(* IEC 61131-3 sources: kns-port-domestic/upstream/plc-process-lib/src/POUs/Devices/FB_AnalogInput, 16 files *)

(* ---- ClassifySignal.method.impl.st ---- *)
IF NOT F_IsFinite(rIn := rIn) THEN
    ClassifySignal := E_AiSignalState.NotFinite;
ELSIF xChannelFault THEN
    ClassifySignal := E_AiSignalState.ChannelFault;
ELSIF stCfgLkg.eInput = E_AiInputType.MilliAmp OR stCfgLkg.eInput = E_AiInputType.Norm420 THEN
    IF stCfgLkg.eInput = E_AiInputType.Norm420 THEN
        rI_mA := GVL_Const.MA_ZERO + GVL_Const.MA_SPAN * rIn;
    ELSE
        rI_mA := rIn;
    END_IF
    IF rI_mA <= GVL_Const.NE43_FAIL_LOW_MA THEN
        ClassifySignal := E_AiSignalState.FailLow;
    ELSIF rI_mA >= GVL_Const.NE43_FAIL_HIGH_MA THEN
        ClassifySignal := E_AiSignalState.FailHigh;
    ELSIF rI_mA < GVL_Const.NE43_MEAS_LOW_MA THEN
        ClassifySignal := E_AiSignalState.UnderRange;
    ELSIF rI_mA > GVL_Const.NE43_MEAS_HIGH_MA THEN
        ClassifySignal := E_AiSignalState.OverRange;
    ELSE
        ClassifySignal := E_AiSignalState.Good;
    END_IF
ELSE
    // Norm01, Eng, Raw: NE 43 не применяется
    ClassifySignal := E_AiSignalState.Good;
END_IF

(* ---- FB_AnalogInput.decl.st ---- *)
// Назначение: аналоговый вход. Сигнал 4–20 мА, нормированный 0–1, инженерные единицы или отсчёты
//             канала → значение в инженерных единицах: достоверность по NAMUR NE 43 с
//             подтверждением tFailDelay и удержанием последнего хорошего значения на время
//             подтверждения, корень с отсечкой малых значений, фильтр первого порядка по реальному
//             шагу времени, уставки HH/H/L/LL (FB_LimitMonitor), подмена значения с ограничением по
//             времени, шесть слотов тревог. Режимы: Auto — измерение, Manual — подмена,
//             OutOfService; Local нет. Наследует FB_DeviceBase: тело — нормативный порядок цикла,
//             шаги обработки сигнала — защищённые методы.
// Автор:      kr0nsch
// Версия:     0.1.0
// Документ:   docs/fb/FB_AnalogInput.md
FUNCTION_BLOCK FB_AnalogInput EXTENDS FB_DeviceBase
VAR_INPUT
    rIn                  : REAL;     // значение канала; смысл — по stCfg.eInput
    xChannelFault        : BOOL;     // диагностика модуля или ошибка обмена (для значений по Modbus)
    xSuppressLimitAlarms : BOOL;     // подавить тревоги уставок по условию (флаги уставок считаются)
END_VAR
VAR_IN_OUT
    stCmd : ST_AnalogInputCmd;       // команды HMI/SCADA (GVL_Hmi.st<TAG>Cmd)
END_VAR
VAR_IN_OUT CONSTANT
    stCfg : ST_AnalogInputCfg;       // параметры (GVL_Persist.st<TAG>Cfg), только чтение
END_VAR
VAR_OUTPUT
    rValue_eu  : REAL;               // значение для логики, инж. ед.
    rValue_pct : REAL;               // значение, % шкалы
    xValid     : BOOL;               // значение пригодно для управления
    xHH        : BOOL;               // верхняя аварийная уставка (после гистерезиса и задержек)
    xH         : BOOL;               // верхняя предупредительная уставка
    xL         : BOOL;               // нижняя предупредительная уставка
    xLL        : BOOL;               // нижняя аварийная уставка
    stSts      : ST_AnalogInputSts;  // состояние для HMI/SCADA
END_VAR
VAR
    stCfgLkg  : ST_AnalogInputCfg;                       // последняя корректная конфигурация (LKG)
    afbLimit  : ARRAY[0..3] OF FB_LimitMonitor;          // уставки, индекс E_AiAlarm.HH, H, L, LL
    fbFail    : FB_Delay;                                // подтверждение отказа сигнала и возврата
    fbOor     : FB_Delay;                                // подтверждение выхода за диапазон и возврата
    fbSubst   : FB_Delay;                                // длительность подмены (tSubstMax)
    eSignal   : E_AiSignalState := E_AiSignalState.Good; // мгновенная классификация сигнала
    xRawFail  : BOOL;                                    // мгновенный отказ сигнала (до подтверждения)
    xFail     : BOOL;                                    // отказ сигнала подтверждён
    xOor      : BOOL;                                    // выход за диапазон подтверждён
    xValueBad : BOOL;                                    // измеренного значения нет: отказ подтверждён
                                                         // или хорошего значения ещё не было
    lrFlt     : LREAL;                                   // состояние фильтра, инж. ед.
    xFltInit  : BOOL := TRUE;                            // фильтр начнётся с текущего значения
    rGood_eu  : REAL;                                    // последнее хорошее значение, инж. ед.
    xHaveGood : BOOL;                                    // хорошее значение было после старта ПЛК или
                                                         // после возврата контроля (OutOfService, Cfg)
    xLowCut   : BOOL;                                    // сработала отсечка малых значений
    xClamped  : BOOL;                                    // значение ограничено шкалой
END_VAR
VAR_TEMP
    eRes       : E_CmdResult;        // результат ProcessMode
    xRawOor    : BOOL;               // мгновенный выход за диапазон (до подтверждения)
    xSupervise : BOOL;               // контроль сигнала: корректная Cfg была, не OutOfService
    xLimOff    : BOOL;               // флаги уставок снять сразу
    xLimSupp   : BOOL;               // подавление тревог уставок
    wLowBits   : WORD;               // младший байт wStatus
    eDevSt     : E_Ne107Status;      // вклад логики устройства в NE 107
END_VAR

(* ---- CallLimit.method.decl.st ---- *)
// Вызов одной уставки FB_LimitMonitor (шаг 7 цикла), результат — флаг уставки xOut. Уставка
// передаётся через VAR_IN_OUT: шаг уставок в теле — один вызов на уставку (AI-1). Внутренний шаг
// устройства: PROTECTED (правило L5 контракта), имя зарезервировано
METHOD PROTECTED CallLimit : BOOL
VAR_INPUT
    rLimValue : REAL;              // контролируемое значение, инж. ед.
    xHigh     : BOOL;              // TRUE — верхняя уставка (HH, H), FALSE — нижняя (L, LL)
    xOff      : BOOL;              // снять флаг сразу (OutOfService, нет Cfg, отказ)
    stLimCfg  : ST_AiLimitCfg;     // параметры уставки (stCfgLkg.astLimit[i])
END_VAR
VAR_IN_OUT
    fbLimit : FB_LimitMonitor;     // уставка afbLimit[i]
END_VAR

(* ---- CheckConfig.method.decl.st ---- *)
// Проверка конфигурации: биты wCfgErr аналогового входа (карта — docs/fb/FB_AnalogInput.md). Только
// считает, ничего не меняет. Сравнения записаны так, чтобы NaN давал ошибку (NOT (x >= a AND x <= b))
METHOD PROTECTED CheckConfig : WORD
VAR_IN_OUT CONSTANT
    stCfgIn : ST_AnalogInputCfg;   // проверяемая конфигурация
END_VAR
VAR
    wErr    : WORD;                // непройденные проверки
    uiIdx   : UINT;                // индекс уставки: HH, H, L, LL
    stLim   : ST_AiLimitCfg;       // копия уставки: короче условия проверок
    xPrev   : BOOL;                // была включённая уставка старше текущей
    rPrevSp : REAL;                // её значение, инж. ед.
    rSpan   : REAL;                // диапазон шкалы, инж. ед.
END_VAR

(* ---- CheckConfig.method.impl.st ---- *)
IF NOT (stCfgIn.eInput = E_AiInputType.MilliAmp OR stCfgIn.eInput = E_AiInputType.Norm420
        OR stCfgIn.eInput = E_AiInputType.Norm01 OR stCfgIn.eInput = E_AiInputType.Eng
        OR stCfgIn.eInput = E_AiInputType.Raw)
THEN
    wErr := wErr OR GVL_Const.AI_CFG_INPUT_TYPE;
END_IF
IF NOT (F_IsFinite(rIn := stCfgIn.rRangeLo_eu) AND F_IsFinite(rIn := stCfgIn.rRangeHi_eu)
        AND stCfgIn.rRangeLo_eu < stCfgIn.rRangeHi_eu)
THEN
    wErr := wErr OR GVL_Const.AI_CFG_RANGE;
END_IF

// Уставки: включённые — в шкале, гистерезис 0 <= h < диапазона, порядок строго LL < L < H < HH
// (обход от HH к LL: каждая следующая включённая строго меньше предыдущей включённой)
rSpan := stCfgIn.rRangeHi_eu - stCfgIn.rRangeLo_eu;
FOR uiIdx := E_AiAlarm.HH TO E_AiAlarm.LL DO
    stLim := stCfgIn.astLimit[uiIdx];
    IF stLim.xEnable THEN
        IF NOT (stLim.rSetpoint_eu >= stCfgIn.rRangeLo_eu AND stLim.rSetpoint_eu <= stCfgIn.rRangeHi_eu) THEN
            wErr := wErr OR GVL_Const.AI_CFG_LIMIT_OUT_OF_RANGE;
        END_IF
        IF NOT (F_IsFinite(rIn := stLim.rHyst_eu) AND stLim.rHyst_eu >= 0.0 AND stLim.rHyst_eu < rSpan) THEN
            wErr := wErr OR GVL_Const.AI_CFG_HYST;
        END_IF
        IF xPrev AND NOT (stLim.rSetpoint_eu < rPrevSp) THEN
            wErr := wErr OR GVL_Const.AI_CFG_LIMIT_ORDER;
        END_IF
        xPrev := TRUE;
        rPrevSp := stLim.rSetpoint_eu;
    END_IF
END_FOR

IF NOT (stCfgIn.rLowCut_pct >= 0.0 AND stCfgIn.rLowCut_pct <= GVL_Const.AI_LOWCUT_MAX_PCT) THEN
    wErr := wErr OR GVL_Const.AI_CFG_LOW_CUT;
END_IF
IF NOT (stCfgIn.eFailValue = E_AiFailValue.HoldLast OR stCfgIn.eFailValue = E_AiFailValue.Substitute)
   OR NOT F_IsFinite(rIn := stCfgIn.rFailValue_eu)
THEN
    wErr := wErr OR GVL_Const.AI_CFG_FAIL_VALUE;
END_IF
IF NOT CheckAlarmCfg(astCfg := stCfgIn.astAlarm) THEN
    wErr := wErr OR GVL_Const.AI_CFG_ALARM;
END_IF
// шкала отсчётов проверяется только у входа Raw: умолчания 0/0 проходят у остальных типов
IF stCfgIn.eInput = E_AiInputType.Raw
   AND NOT (F_IsFinite(rIn := stCfgIn.rRawLo_cnt) AND F_IsFinite(rIn := stCfgIn.rRawHi_cnt)
            AND stCfgIn.rRawLo_cnt < stCfgIn.rRawHi_cnt)
THEN
    wErr := wErr OR GVL_Const.AI_CFG_RAW_RANGE;
END_IF
CheckConfig := wErr;

(* ---- ClassifySignal.method.decl.st ---- *)
// Шаг 6.1 цикла: мгновенная классификация сигнала (до подтверждения tFailDelay). NE 43 — только для
// MilliAmp и Norm420 (I = 4 + 16·rIn); старшинство NotFinite > ChannelFault > FailLow/FailHigh >
// UnderRange/OverRange > Good. Границы 3,6 и 21,0 мА включены в отказ (A-02, сверить с NAMUR NE 43).
// Читает входы rIn, xChannelFault и stCfgLkg; ничего не меняет
METHOD PROTECTED ClassifySignal : E_AiSignalState
VAR
    rI_mA : REAL;   // ток для проверки NE 43, мА
END_VAR

(* ---- ComputeValue.method.decl.st ---- *)
// Шаг 6.3 цикла (LREAL): нормировка по типу входа, корень и отсечка малых значений, инженерные
// единицы, ограничение шкалой, фильтр первого порядка — точная экспонента по реальному шагу времени.
// 4–20 мА (MilliAmp, Norm420): значение не экстраполируется за насыщение NE 43 (3,8 и 20,5 мА, AI-13)
// ltDt (реакция не зависит от цикла). Без расчёта (xCompute = FALSE: нет корректной Cfg, OutOfService,
// отказ сигнала) фильтр стоит. После подтверждённого отказа и после возврата контроля (xRestart) фильтр
// начинается с текущего значения, без «подтягивания» от старого; короткий неподтверждённый провал
// фильтр только замораживает — после него значение продолжается без скачка (AI-12). Хорошее значение
// для удержания запоминается, пока отказ не подтверждён
METHOD PROTECTED ComputeValue
VAR_INPUT
    xCompute : BOOL;   // значение считается в этом вызове
    xRestart : BOOL;   // фильтр начать заново: отказ подтверждён или сигнал не контролируется
END_VAR
VAR
    lrLo   : LREAL;    // начало шкалы, инж. ед.
    lrSpan : LREAL;    // диапазон шкалы, инж. ед.
    lrX    : LREAL;    // нормированное значение, доли шкалы
    lrEng  : LREAL;    // значение до фильтра, инж. ед.
    lrT_s  : LREAL;    // постоянная времени фильтра, с
    lrSane : LREAL;    // предел |значения| REAL_SANE_MAX
    lrXLo  : LREAL;    // насыщение NE 43 снизу (3,8 мА), доли шкалы
    lrXHi  : LREAL;    // насыщение NE 43 сверху (20,5 мА), доли шкалы
END_VAR

(* ---- ComputeValue.method.impl.st ---- *)
xLowCut := FALSE;
xClamped := FALSE;
IF xCompute THEN
    // нормировка: x — доли шкалы
    lrLo := REAL_TO_LREAL(stCfgLkg.rRangeLo_eu);
    lrSpan := REAL_TO_LREAL(stCfgLkg.rRangeHi_eu) - lrLo;
    IF stCfgLkg.eInput = E_AiInputType.MilliAmp THEN
        lrX := (REAL_TO_LREAL(rIn) - REAL_TO_LREAL(GVL_Const.MA_ZERO)) / REAL_TO_LREAL(GVL_Const.MA_SPAN);
    ELSIF stCfgLkg.eInput = E_AiInputType.Eng THEN
        lrX := (REAL_TO_LREAL(rIn) - lrLo) / lrSpan;
    ELSIF stCfgLkg.eInput = E_AiInputType.Raw THEN
        lrX := (REAL_TO_LREAL(rIn) - REAL_TO_LREAL(stCfgLkg.rRawLo_cnt))
               / (REAL_TO_LREAL(stCfgLkg.rRawHi_cnt) - REAL_TO_LREAL(stCfgLkg.rRawLo_cnt));
    ELSE
        // Norm420, Norm01: вход уже в долях шкалы
        lrX := REAL_TO_LREAL(rIn);
    END_IF
    // NE 43: за насыщением 3,8 / 20,5 мА измерения нет — это защитные полосы до порогов отказа (ток отказа с
    // погрешностью канала или насыщение датчика). Значение не экстраполируется дальше насыщения (AI-13)
    IF stCfgLkg.eInput = E_AiInputType.MilliAmp OR stCfgLkg.eInput = E_AiInputType.Norm420 THEN
        lrXLo := (REAL_TO_LREAL(GVL_Const.NE43_MEAS_LOW_MA) - REAL_TO_LREAL(GVL_Const.MA_ZERO))
                 / REAL_TO_LREAL(GVL_Const.MA_SPAN);
        lrXHi := (REAL_TO_LREAL(GVL_Const.NE43_MEAS_HIGH_MA) - REAL_TO_LREAL(GVL_Const.MA_ZERO))
                 / REAL_TO_LREAL(GVL_Const.MA_SPAN);
        lrX := LIMIT(lrXLo, lrX, lrXHi);
    END_IF

    // корень (расход по перепаду давления), затем отсечка — она действует и без корня
    IF stCfgLkg.xSqrt THEN
        lrX := SQRT(MAX(lrX, 0.0));
    END_IF
    IF stCfgLkg.rLowCut_pct > 0.0
       AND lrX * REAL_TO_LREAL(GVL_Const.PCT_FULL) < REAL_TO_LREAL(stCfgLkg.rLowCut_pct)
    THEN
        lrX := 0.0;
        xLowCut := TRUE;
    END_IF

    // инженерные единицы; по умолчанию — экстраполяция за шкалу, при xClamp — ограничение шкалой
    lrEng := lrLo + lrX * lrSpan;
    IF stCfgLkg.xClamp THEN
        IF lrEng < lrLo THEN
            lrEng := lrLo;
            xClamped := TRUE;
        ELSIF lrEng > lrLo + lrSpan THEN
            lrEng := lrLo + lrSpan;
            xClamped := TRUE;
        END_IF
    END_IF

    // фильтр: alpha = 1 - exp(-dt / T); T#0S, первый расчёт и расчёт после подтверждённого отказа — без фильтра
    lrT_s := F_TimeToSec(tIn := stCfgLkg.tFilter);
    IF xFltInit OR lrT_s <= 0.0 THEN
        lrFlt := lrEng;
    ELSE
        lrFlt := lrFlt + (1.0 - EXP(-F_LTimeToSec(ltIn := ltDt) / lrT_s)) * (lrEng - lrFlt);
    END_IF
    xFltInit := FALSE;

    // хорошее значение для удержания: пока отказ не подтверждён; |значение| не больше REAL_SANE_MAX
    IF NOT xFail THEN
        lrSane := REAL_TO_LREAL(GVL_Const.REAL_SANE_MAX);
        rGood_eu := LREAL_TO_REAL(LIMIT(-lrSane, lrFlt, lrSane));
        xHaveGood := TRUE;
    END_IF
ELSE
    // расчёта нет. Отказ подтверждён или сигнал не контролируется (xRestart): фильтр начнётся заново с
    // текущего значения. Неподтверждённый провал фильтр замораживает: после него — продолжение без скачка
    xFltInit := xFltInit OR xRestart;
END_IF

(* ---- FaultBits.method.impl.st ---- *)
IF xFail AND eSignal = E_AiSignalState.FailLow THEN
    FaultBits := GVL_Const.AI_FLT_FAIL_LOW;
ELSIF xFail AND eSignal = E_AiSignalState.FailHigh THEN
    FaultBits := GVL_Const.AI_FLT_FAIL_HIGH;
ELSIF xFail AND eSignal = E_AiSignalState.ChannelFault THEN
    FaultBits := GVL_Const.AI_FLT_CHANNEL;
ELSIF xFail AND eSignal = E_AiSignalState.NotFinite THEN
    FaultBits := GVL_Const.AI_FLT_NOT_FINITE;
ELSE
    // отказа нет или сигнал уже вернулся (идёт подтверждение возврата)
    FaultBits := 0;
END_IF

(* ---- FB_AnalogInput.impl.st ---- *)
// 0. Первый вызов (до ProcessMode): тип, число слотов тревог; режим «Измерение» в памяти режима,
//    подмена (Manual) даёт CheckFunction
IF xFirstCall THEN
    uiAlarmCount := GVL_Const.AI_ALARM_COUNT;
    eDevType := E_DeviceType.AnalogInput;
    xManualIsCheck := TRUE;
    stModeMem.eRemoteMode := E_DeviceMode.Auto;
END_IF

// 1. Время
BeginCycle();

// 2. Конфигурация (LKG): дальше логика читает только stCfgLkg
IF AcceptCfg(wErr := CheckConfig(stCfgIn := stCfg)) THEN
    stCfgLkg := stCfg;
END_IF

// 3. Reset: фиксируемых отказов нет (отказ сигнала снимается сам), результат команды — Accepted;
//    квитирование выполнит RunAlarms
IF xResetReq OR stCmd.stCommon.xReset THEN
    SetCmdResult(eResult := E_CmdResult.Accepted);
END_IF

// 4. Режим: Local нет, OutOfService разрешён всегда; память режима — stModeMem (подмена и вывод из
//    работы не переживают перезапуск ПЛК, A-06)
eRes := ProcessMode(xLocalSel := FALSE, xLocalSupported := FALSE, xOosAllowed := TRUE,
                    stCmd := stCmd.stCommon, stRetain := stModeMem);
IF eRes <> E_CmdResult.None THEN
    SetCmdResult(eResult := eRes);
END_IF

// 5. Подмена ограничена по времени: Manual длится tSubstMax — возврат в Auto (SubstExpired). До выбора
//    значения: в этом же вызове значение уже измеренное. Preset — чтобы новый запрос подмены в
//    следующем вызове отсчитал tSubstMax заново
fbSubst(xIn := (eMode = E_DeviceMode.Manual) AND (stCfgLkg.tSubstMax > T#0S), tOnDelay := stCfgLkg.tSubstMax,
        itfTime := itfTimeAct);
IF fbSubst.xOut THEN
    SwitchRemoteMode(eNew := E_DeviceMode.Auto, stRetain := stModeMem);
    fbSubst.Preset(xValue := FALSE);
    SetCmdResult(eResult := E_CmdResult.SubstExpired);
END_IF

// 6. Сигнал и значение
// 6.1 Классификация (мгновенная, NE 43)
eSignal := ClassifySignal();
xRawFail := eSignal = E_AiSignalState.NotFinite OR eSignal = E_AiSignalState.ChannelFault
            OR eSignal = E_AiSignalState.FailLow OR eSignal = E_AiSignalState.FailHigh;
xRawOor := eSignal = E_AiSignalState.UnderRange OR eSignal = E_AiSignalState.OverRange;
// 6.2 Подтверждение: и появление, и возврат — через tFailDelay. Без корректной Cfg (тип входа ещё не
//     известен) и в OutOfService сигнал не контролируется: флаги снимаются сразу, отсчёт — заново.
//     Последнее хорошее значение при этом устаревает (датчик могли сменить «в ремонте»): после возврата
//     контроля удерживать нечего, как после старта ПЛК (AI-2)
xSupervise := xCfgEverOk AND eMode <> E_DeviceMode.OutOfService;
IF xSupervise THEN
    fbFail(xIn := xRawFail, tOnDelay := stCfgLkg.tFailDelay, tOffDelay := stCfgLkg.tFailDelay,
           itfTime := itfTimeAct);
    fbOor(xIn := xRawOor AND NOT xRawFail, tOnDelay := stCfgLkg.tFailDelay, tOffDelay := stCfgLkg.tFailDelay,
          itfTime := itfTimeAct);
ELSE
    fbFail.Preset(xValue := FALSE);
    fbOor.Preset(xValue := FALSE);
    xHaveGood := FALSE;
END_IF
xFail := fbFail.xOut;
xOor := fbOor.xOut;
// 6.3 Значение и фильтр: не считаются без корректной Cfg, в OutOfService и пока сигнал отказал. Фильтр
//     начинается заново после подтверждённого отказа и после возврата контроля; короткий провал его только
//     замораживает (AI-12)
ComputeValue(xCompute := xSupervise AND NOT xRawFail, xRestart := xFail OR NOT xSupervise);
// 6.4 Выбор значения по режиму и состоянию сигнала
xValueBad := xFail OR (xRawFail AND NOT xHaveGood);
SelectValue(rSubst_eu := stCmd.rSubstValue_eu);

// 7. Уставки — по выбранному значению (в Manual — по подменённому: так при наладке проверяют
//    блокировки). Флаги снимаются сразу в OutOfService, без корректной Cfg и в Auto без измеренного
//    значения, если не xLimitsOnFail
xLimOff := eMode = E_DeviceMode.OutOfService OR NOT xCfgEverOk
           OR (eMode = E_DeviceMode.Auto AND xValueBad AND NOT stCfgLkg.xLimitsOnFail);
xHH := CallLimit(rLimValue := rValue_eu, xHigh := TRUE, xOff := xLimOff,
                 stLimCfg := stCfgLkg.astLimit[E_AiAlarm.HH], fbLimit := afbLimit[E_AiAlarm.HH]);
xH := CallLimit(rLimValue := rValue_eu, xHigh := TRUE, xOff := xLimOff,
                stLimCfg := stCfgLkg.astLimit[E_AiAlarm.H], fbLimit := afbLimit[E_AiAlarm.H]);
xL := CallLimit(rLimValue := rValue_eu, xHigh := FALSE, xOff := xLimOff,
                stLimCfg := stCfgLkg.astLimit[E_AiAlarm.L], fbLimit := afbLimit[E_AiAlarm.L]);
xLL := CallLimit(rLimValue := rValue_eu, xHigh := FALSE, xOff := xLimOff,
                 stLimCfg := stCfgLkg.astLimit[E_AiAlarm.LL], fbLimit := afbLimit[E_AiAlarm.LL]);

// 8. Слежение: пока значением управляет не оператор, ФБ пишет текущее значение в поле подмены —
//    переход в подмену без рывка
IF eMode <> E_DeviceMode.Manual THEN
    stCmd.rSubstValue_eu := rValue_eu;
END_IF

// 9. Тревоги (слоты E_AiAlarm). Значение события: rValue_eu, у слота Failure — сырое rIn
xLimSupp := xSuppressLimitAlarms OR (xFail AND NOT stCfgLkg.xLimitsOnFail);
axAlmCond[E_AiAlarm.HH] := xHH;
axAlmCond[E_AiAlarm.H] := xH;
axAlmCond[E_AiAlarm.L] := xL;
axAlmCond[E_AiAlarm.LL] := xLL;
axAlmCond[E_AiAlarm.Failure] := xFail;
axAlmCond[E_AiAlarm.OutOfRange] := xOor AND NOT xFail;
axAlmSuppress[E_AiAlarm.HH] := xLimSupp;
axAlmSuppress[E_AiAlarm.H] := xLimSupp;
axAlmSuppress[E_AiAlarm.L] := xLimSupp;
axAlmSuppress[E_AiAlarm.LL] := xLimSupp;
axAlmSuppress[E_AiAlarm.Failure] := FALSE;
axAlmSuppress[E_AiAlarm.OutOfRange] := FALSE;
arAlmValue[E_AiAlarm.HH] := rValue_eu;
arAlmValue[E_AiAlarm.H] := rValue_eu;
arAlmValue[E_AiAlarm.L] := rValue_eu;
arAlmValue[E_AiAlarm.LL] := rValue_eu;
arAlmValue[E_AiAlarm.Failure] := rIn;
arAlmValue[E_AiAlarm.OutOfRange] := rValue_eu;
RunAlarms(udiIdBase := stCfgLkg.udiAlarmIdBase, stCmd := stCmd.stCommon, astCfg := stCfgLkg.astAlarm);

// 10. Состояние. AI_STS_FAIL_PENDING — в Auto последнее хорошее значение удерживается как годное до
//     подтверждения отказа (не при xValueBad: удерживать нечего, AI-2)
wLowBits := SEL(xHH, 0, GVL_Const.AI_STS_HH) OR SEL(xH, 0, GVL_Const.AI_STS_H)
            OR SEL(xL, 0, GVL_Const.AI_STS_L) OR SEL(xLL, 0, GVL_Const.AI_STS_LL)
            OR SEL(xFail, 0, GVL_Const.AI_STS_SIGNAL_FAIL) OR SEL(xOor, 0, GVL_Const.AI_STS_OUT_OF_RANGE)
            OR SEL(eMode = E_DeviceMode.Auto AND xSupervise AND xRawFail AND NOT xValueBad, 0,
                   GVL_Const.AI_STS_FAIL_PENDING)
            OR SEL(xLowCut, 0, GVL_Const.AI_STS_LOW_CUT);
IF xFail THEN
    eDevSt := E_Ne107Status.Failure;
ELSIF xOor THEN
    eDevSt := E_Ne107Status.OutOfSpecification;
ELSE
    eDevSt := E_Ne107Status.Good;
END_IF
stSts.rValue_eu := rValue_eu;
stSts.rValue_pct := rValue_pct;
stSts.rIn := rIn;
stSts.eSignal := eSignal;
stSts.uiSubstRemain_s := SubstRemainSec();
FinishCycle(eDevStatus := eDevSt, xAvailableDev := xValid, wLow := wLowBits, wFaultBits := FaultBits(),
            wWarnBits := WarningBits(), stCommon := stSts.stCommon);

(* ---- SelectValue.method.decl.st ---- *)
// Шаг 6.4 цикла: значение для логики rValue_eu, rValue_pct и xValid по режиму и состоянию сигнала
// (таблица 11.3 контракта). Удержание последнего хорошего значения на время подтверждения отказа:
// обрыв не даёт мгновенного ложного LL. Если хорошего значения после старта ПЛК или после выхода
// из OutOfService ещё не было (xValueBad при неподтверждённом отказе), удерживать нечего — значение
// как при подтверждённом отказе, xValid = FALSE (AI-2). Выход за диапазон NE 43 подтверждён (xOor) —
// значение насыщения (граница, процесс за ней неизвестен), xValid = FALSE (AI-13). Значение подмены приходит
// параметром: метод не читает VAR_IN_OUT (R2)
METHOD PROTECTED SelectValue
VAR_INPUT
    rSubst_eu : REAL;   // значение подмены stCmd.rSubstValue_eu, инж. ед.
END_VAR
VAR
    lrSane : LREAL;     // предел |значения| REAL_SANE_MAX
END_VAR

(* ---- SelectValue.method.impl.st ---- *)
IF NOT xCfgEverOk THEN
    // безопасное значение: корректной Cfg ещё не было
    rValue_eu := 0.0;
    xValid := FALSE;
ELSIF eMode = E_DeviceMode.OutOfService THEN
    // значение удерживается
    xValid := FALSE;
ELSIF eMode = E_DeviceMode.Manual THEN
    // подмена без фильтра; неконечное значение подмены не принимается (значение удерживается)
    IF F_IsFinite(rIn := rSubst_eu) THEN
        rValue_eu := rSubst_eu;
    END_IF
    xValid := TRUE;
ELSIF xValueBad THEN
    IF stCfgLkg.eFailValue = E_AiFailValue.Substitute THEN
        rValue_eu := stCfgLkg.rFailValue_eu;
    ELSE
        rValue_eu := rGood_eu;
    END_IF
    xValid := FALSE;
ELSE
    // хорошее значение, значение насыщения NE 43 или последнее хорошее до подтверждения отказа
    // (AI_STS_FAIL_PENDING). Подтверждённый выход за диапазон — для управления непригодно (AI-13): ПИД и
    // автоматика не работают по значению, за которым процесс неизвестен (ток отказа NAMUR, прочитанный с
    // погрешностью канала, тоже попадает в защитную полосу); уставки по нему считаются
    rValue_eu := rGood_eu;
    xValid := NOT xOor;
END_IF

IF xCfgEverOk THEN
    lrSane := REAL_TO_LREAL(GVL_Const.REAL_SANE_MAX);
    rValue_pct := LREAL_TO_REAL(LIMIT(-lrSane,
                                      (REAL_TO_LREAL(rValue_eu) - REAL_TO_LREAL(stCfgLkg.rRangeLo_eu))
                                      / (REAL_TO_LREAL(stCfgLkg.rRangeHi_eu) - REAL_TO_LREAL(stCfgLkg.rRangeLo_eu))
                                      * REAL_TO_LREAL(GVL_Const.PCT_FULL),
                                      lrSane));
ELSE
    rValue_pct := 0.0;
END_IF

(* ---- SubstRemainSec.method.decl.st ---- *)
// Остаток подмены для stSts.uiSubstRemain_s: целые секунды с округлением вверх (пока подмена идёт,
// остаток не 0), не больше UINT_MAX. 0 — подмены нет или её срок не ограничен (tSubstMax = T#0S)
METHOD PROTECTED SubstRemainSec : UINT
VAR
    lrRemain_s  : LREAL;   // до снятия подмены, с
    udiRemain_s : UDINT;   // то же, целых секунд
END_VAR

(* ---- SubstRemainSec.method.impl.st ---- *)
IF eMode = E_DeviceMode.Manual AND stCfgLkg.tSubstMax > T#0S THEN
    lrRemain_s := F_TimeToSec(tIn := fbSubst.tRemaining);
    udiRemain_s := LREAL_TO_UDINT(lrRemain_s);
    IF UDINT_TO_LREAL(udiRemain_s) < lrRemain_s THEN
        udiRemain_s := udiRemain_s + 1;
    END_IF
    SubstRemainSec := UDINT_TO_UINT(MIN(udiRemain_s, UINT_TO_UDINT(GVL_Const.UINT_MAX)));
ELSE
    SubstRemainSec := 0;
END_IF

(* ---- WarningBits.method.decl.st ---- *)
// Слово wWarning: пока выход за диапазон подтверждён (xOor) — бит по текущей классификации;
// AI_WRN_CLAMPED — значение этого вызова ограничено шкалой (контракт 11.5)
METHOD PROTECTED WarningBits : WORD
VAR
    wBits : WORD;   // собранные биты
END_VAR

(* ---- WarningBits.method.impl.st ---- *)
IF xOor AND eSignal = E_AiSignalState.UnderRange THEN
    wBits := GVL_Const.AI_WRN_UNDER_RANGE;
ELSIF xOor AND eSignal = E_AiSignalState.OverRange THEN
    wBits := GVL_Const.AI_WRN_OVER_RANGE;
END_IF
IF xClamped THEN
    wBits := wBits OR GVL_Const.AI_WRN_CLAMPED;
END_IF
WarningBits := wBits;
